// TIA Portal V18 export
TYPE "UserValidationMdz_in"
   STRUCT
      Station : Array[1.."Station_Setup_Const"] of Struct
         UserMaster_ID : DInt;
         Position_ID_Validation : Int;
         LogIn : Bool;
         Position : Array[1.."Position_Setup_Const"] of Struct
            User_ID : DInt;
            BadgeNumber : LInt;
            LogIn : Bool;
            LogOut : Bool;
            ByPass : Bool;
         END_STRUCT;
      END_STRUCT;
   END_STRUCT;
   // Station[1..20].UserMaster_ID := 0;
   // Station[1..20].Position_ID_Validation := 0;
   // Station[1..20].LogIn := FALSE;
   // Station[1].Position[1].User_ID := 0;
   // Station[2].Position[1].User_ID := 0;
   // Station[3].Position[1].User_ID := 0;
   // Station[4].Position[1].User_ID := 0;
   // Station[5].Position[1].User_ID := 0;
   // Station[6].Position[1].User_ID := 0;
   // Station[7].Position[1].User_ID := 0;
   // Station[8].Position[1].User_ID := 0;
   // Station[9].Position[1].User_ID := 0;
   // Station[10].Position[1].User_ID := 0;
   // Station[11].Position[1].User_ID := 0;
   // Station[12].Position[1].User_ID := 0;
   // Station[13].Position[1].User_ID := 0;
   // Station[14].Position[1].User_ID := 0;
   // Station[15].Position[1].User_ID := 0;
   // Station[16].Position[1].User_ID := 0;
   // Station[17].Position[1].User_ID := 0;
   // Station[18].Position[1].User_ID := 0;
   // Station[19].Position[1].User_ID := 0;
   // Station[20].Position[1].User_ID := 0;
   // Station[1].Position[1].BadgeNumber := 0;
   // Station[2].Position[1].BadgeNumber := 0;
   // Station[3].Position[1].BadgeNumber := 0;
   // Station[4].Position[1].BadgeNumber := 0;
   // Station[5].Position[1].BadgeNumber := 0;
   // Station[6].Position[1].BadgeNumber := 0;
   // Station[7].Position[1].BadgeNumber := 0;
   // Station[8].Position[1].BadgeNumber := 0;
   // Station[9].Position[1].BadgeNumber := 0;
   // Station[10].Position[1].BadgeNumber := 0;
   // Station[11].Position[1].BadgeNumber := 0;
   // Station[12].Position[1].BadgeNumber := 0;
   // Station[13].Position[1].BadgeNumber := 0;
   // Station[14].Position[1].BadgeNumber := 0;
   // Station[15].Position[1].BadgeNumber := 0;
   // Station[16].Position[1].BadgeNumber := 0;
   // Station[17].Position[1].BadgeNumber := 0;
   // Station[18].Position[1].BadgeNumber := 0;
   // Station[19].Position[1].BadgeNumber := 0;
   // Station[20].Position[1].BadgeNumber := 0;
   // Station[1].Position[1].LogIn := FALSE;
   // Station[2].Position[1].LogIn := FALSE;
   // Station[3].Position[1].LogIn := FALSE;
   // Station[4].Position[1].LogIn := FALSE;
   // Station[5].Position[1].LogIn := FALSE;
   // Station[6].Position[1].LogIn := FALSE;
   // Station[7].Position[1].LogIn := FALSE;
   // Station[8].Position[1].LogIn := FALSE;
   // Station[9].Position[1].LogIn := FALSE;
   // Station[10].Position[1].LogIn := FALSE;
   // Station[11].Position[1].LogIn := FALSE;
   // Station[12].Position[1].LogIn := FALSE;
   // Station[13].Position[1].LogIn := FALSE;
   // Station[14].Position[1].LogIn := FALSE;
   // Station[15].Position[1].LogIn := FALSE;
   // Station[16].Position[1].LogIn := FALSE;
   // Station[17].Position[1].LogIn := FALSE;
   // Station[18].Position[1].LogIn := FALSE;
   // Station[19].Position[1].LogIn := FALSE;
   // Station[20].Position[1].LogIn := FALSE;
   // Station[1].Position[1].LogOut := TRUE;
   // Station[2].Position[1].LogOut := TRUE;
   // Station[3].Position[1].LogOut := TRUE;
   // Station[4].Position[1].LogOut := TRUE;
   // Station[5].Position[1].LogOut := TRUE;
   // Station[6].Position[1].LogOut := TRUE;
   // Station[7].Position[1].LogOut := TRUE;
   // Station[8].Position[1].LogOut := TRUE;
   // Station[9].Position[1].LogOut := TRUE;
   // Station[10].Position[1].LogOut := TRUE;
   // Station[11].Position[1].LogOut := TRUE;
   // Station[12].Position[1].LogOut := TRUE;
   // Station[13].Position[1].LogOut := TRUE;
   // Station[14].Position[1].LogOut := TRUE;
   // Station[15].Position[1].LogOut := TRUE;
   // Station[16].Position[1].LogOut := TRUE;
   // Station[17].Position[1].LogOut := TRUE;
   // Station[18].Position[1].LogOut := TRUE;
   // Station[19].Position[1].LogOut := TRUE;
   // Station[20].Position[1].LogOut := TRUE;
   // Station[1].Position[1].ByPass := FALSE;
   // Station[2].Position[1].ByPass := FALSE;
   // Station[3].Position[1].ByPass := FALSE;
   // Station[4].Position[1].ByPass := FALSE;
   // Station[5].Position[1].ByPass := FALSE;
   // Station[6].Position[1].ByPass := FALSE;
   // Station[7].Position[1].ByPass := FALSE;
   // Station[8].Position[1].ByPass := FALSE;
   // Station[9].Position[1].ByPass := FALSE;
   // Station[10].Position[1].ByPass := FALSE;
   // Station[11].Position[1].ByPass := FALSE;
   // Station[12].Position[1].ByPass := FALSE;
   // Station[13].Position[1].ByPass := FALSE;
   // Station[14].Position[1].ByPass := FALSE;
   // Station[15].Position[1].ByPass := FALSE;
   // Station[16].Position[1].ByPass := FALSE;
   // Station[17].Position[1].ByPass := FALSE;
   // Station[18].Position[1].ByPass := FALSE;
   // Station[19].Position[1].ByPass := FALSE;
   // Station[20].Position[1].ByPass := FALSE;
END_TYPE
